Yaskawa INFORM job: MANYMOV.JBI

/JOB
//NAME MANYMOV
//POS
///NPOS 40,0,0,0,0,0
///TOOL 9
///POSTYPE PULSE
///PULSE
C00000=0,-10240,0,-34475,0,0,22983
C00001=0,-10240,0,-34475,0,0,22983
C00002=20480,-10240,0,-34475,0,-8704,22983
C00003=0,-10240,0,-34475,0,0,22983
C00004=0,-10240,0,-34475,0,0,22983
C00005=0,-10240,0,-34475,0,0,22983
C00006=20480,-10240,0,-34475,0,-8704,22983
C00007=0,-10240,0,-34475,0,0,22983
C00008=0,-10240,0,-34475,0,0,22983
C00009=0,-10240,0,-34475,0,0,22983
C00010=20480,-10240,0,-34475,0,-8704,22983
C00011=0,-10240,0,-34475,0,0,22983
C00012=0,-10240,0,-34475,0,0,22983
C00013=0,-10240,0,-34475,0,0,22983
C00014=20480,-10240,0,-34475,0,-8704,22983
C00015=0,-10240,0,-34475,0,0,22983
C00016=0,-10240,0,-34475,0,0,22983
C00017=0,-10240,0,-34475,0,0,22983
C00018=20480,-10240,0,-34475,0,-8704,22983
C00019=0,-10240,0,-34475,0,0,22983
C00020=0,-10240,0,-34475,0,0,22983
C00021=0,-10240,0,-34475,0,0,22983
C00022=20480,-10240,0,-34475,0,-8704,22983
C00023=0,-10240,0,-34475,0,0,22983
C00024=0,-10240,0,-34475,0,0,22983
C00025=0,-10240,0,-34475,0,0,22983
C00026=20480,-10240,0,-34475,0,-8704,22983
C00027=0,-10240,0,-34475,0,0,22983
C00028=0,-10240,0,-34475,0,0,22983
C00029=0,-10240,0,-34475,0,0,22983
C00030=20480,-10240,0,-34475,0,-8704,22983
C00031=0,-10240,0,-34475,0,0,22983
C00032=0,-10240,0,-34475,0,0,22983
C00033=0,-10240,0,-34475,0,0,22983
C00034=20480,-10240,0,-34475,0,-8704,22983
C00035=0,-10240,0,-34475,0,0,22983
C00036=0,-10240,0,-34475,0,0,22983
C00037=0,-10240,0,-34475,0,0,22983
C00038=20480,-10240,0,-34475,0,-8704,22983
C00039=0,-10240,0,-34475,0,0,22983
//INST
<volatile>
///COMM Generated using RoboDK
///ATTR SC,RW
///GROUP1 RB1
NOP
'Program generated by RoboDK v
'6.0.7 for Yaskawa Motoman CSD
'A10F on XX/XX/XXXX 18:00:00
'Using nominal kinematics.
'Using Frame S (targets wrt ba
'se):
'1234.6,-98.8,50.5,0.0,0.0,30.
'0
'Tool Tool S should be close t
'o:
'10.0,20.0,150.0,0.0,0.0,0.0
MOVJ C00000 VJ=50.00
MOVL C00001 V=500.0
MOVJ C00002 VJ=50.00
MOVL C00003 V=500.0
MOVJ C00004 VJ=50.00
MOVL C00005 V=500.0
MOVJ C00006 VJ=50.00
MOVL C00007 V=500.0
MOVJ C00008 VJ=50.00
MOVL C00009 V=500.0
MOVJ C00010 VJ=50.00
MOVL C00011 V=500.0
MOVJ C00012 VJ=50.00
MOVL C00013 V=500.0
MOVJ C00014 VJ=50.00
MOVL C00015 V=500.0
MOVJ C00016 VJ=50.00
MOVL C00017 V=500.0
MOVJ C00018 VJ=50.00
MOVL C00019 V=500.0
MOVJ C00020 VJ=50.00
MOVL C00021 V=500.0
MOVJ C00022 VJ=50.00
MOVL C00023 V=500.0
MOVJ C00024 VJ=50.00
MOVL C00025 V=500.0
MOVJ C00026 VJ=50.00
MOVL C00027 V=500.0
MOVJ C00028 VJ=50.00
MOVL C00029 V=500.0
MOVJ C00030 VJ=50.00
MOVL C00031 V=500.0
MOVJ C00032 VJ=50.00
MOVL C00033 V=500.0
MOVJ C00034 VJ=50.00
MOVL C00035 V=500.0
MOVJ C00036 VJ=50.00
MOVL C00037 V=500.0
MOVJ C00038 VJ=50.00
MOVL C00039 V=500.0
END
